FUNCTION_BLOCK FB_ModeSelect
VAR_INPUT
	bInterlockBypass: BOOL;
	bAutoPlayEnable: BOOL:=TRUE;
	sModuleDescription: STRING:='Mode Select';
	eModeZone:E_ModeZone;
	bLockedFB: BOOL;
	bPistonCheck: BOOL:=TRUE;
	bStateSafe_mode: BOOL:=TRUE;
END_VAR
VAR_OUTPUT
	bModeStillState: BOOL;
	bLockRequest: BOOL;
END_VAR
VAR
	fbPrintErrMessageByID: FB_PrintErrMessageByID_SFC_Cycle;
	r_trig_ModeExchange1: R_TRIG;
	r_trig_ModeExchange2: R_TRIG;
	r_trig_ModeExchange3: R_TRIG;
	ton_ModeExchengeDelay: TON;	
	fbOperation:FB_Operation;
	bLockRelay: BOOL;	
	i: INT;
	bPistonsOK: BOOL;
	fbFormatString:FB_FormatString;
	sFB_ID: STRING(3):='050';

	sActErrorID: STRING(11);
	sFullErrorId: STRING(11);
	//r_trigAuto: R_TRIG;
	r_trigIntClose: R_TRIG;
	r_trigIntOpen: R_TRIG;
	bIntZonePaused: BOOL;
	rt_Play: R_TRIG;

END_VAR
VAR
	ton_ResumeMachine: TON;
	ton_ResetErrors: TON;
	ton_ResetAllCycles: TON;
	ton_PlayAllDelay: TON;
	ton_PauseDelay: TON;
	r_trigPlayAllDelay: R_TRIG;
	ton_PlayDelay: TON;
END_VAR
VAR_IN_OUT
	stMode:ST_Mode;
	stOperation:ST_OperationButtons;
END_VAR

act_Oper();
act_ModeStillState();
fbOperation(stOper:=stOperation);
stMode.eModeZone:=eModeZone;		
stOperation.eModeZone:=eModeZone;
stOperation.sModeZone:=TO_STRING(eModeZone);
IF (stMode.iActMode=E_WorkingMode.eAutoMode OR stMode.iActMode=E_WorkingMode.eSemiAutoMode)
AND NOT bInterlockBypass
THEN;
	bLockRequest:=TRUE;
ELSE;
	bLockRequest:=FALSE;
END_IF



r_trigIntClose(CLK:=bLockedFB);
r_trigIntOpen(CLK:=NOT bLockedFB);

(*888888888888888888   InterLocks Zone 1		8888888888888*)
IF stOperation.iActOperation=E_OperationButtons.ePlayAll AND  r_trigIntOpen.Q THEN
	bIntZonePaused:=TRUE;
END_IF

IF NOT bLockedFB 
AND NOT bInterlockBypass	
AND stOperation.iActOperation=E_OperationButtons.ePlayAll THEN
	//Message
	sActErrorID:='351'; // '050x000x351',	'Warning',	'Interlock Paused Operation',
	act_GetErrorID_Format();
	fbPrintErrMessageByID(sFB_ModuleDescription:=sModuleDescription,sActErrorID:=sFullErrorId,bSFCError:=TRUE);
	stOperation.bSetPause:=TRUE;
	stOperation.iPauseHistory:=4;
END_IF


IF bAutoPlayEnable AND bIntZonePaused AND r_trigIntClose.Q THEN
	stOperation.bSetPlay:=TRUE;
	bIntZonePaused:=FALSE;
END_IF

IF bLockedFB OR stMode.iActMode=E_WorkingMode.eManualMode THEN
	bIntZonePaused:=FALSE;
END_IF

rt_Play(CLK:=stOperation.iActOperation=E_OperationButtons.ePlayAll);

IF NOT bStateSafe_mode OR stOperation.bStopResetAll THEN;
	stMode.bSetManual:=TRUE;
	stOperation.bSetPause:=TRUE;
END_IF

stMode.bStateSafe_mode:=stOperation.bStateSafe_mode:=bStateSafe_mode;

m_Error_zone_check();

stOperation.iActModeState:=stMode.iActMode;

ACTION act_AutomationLock_Failed:
sActErrorID:='306';//'050x000x306',	'Warning',	'Semi/Auto mode request rejected, automation lock failed',
act_GetErrorID_Format();
fbPrintErrMessageByID(sFB_ModuleDescription:=sModuleDescription,sActErrorID:=sFullErrorId,bSFCError:=TRUE);
END_ACTION

ACTION act_Done:
stMode.bSetManual:=FALSE;
stMode.bSetSemi:=FALSE;
stMode.bSetAuto:=FALSE;
//stMode.iErrorNum:=0;
//stMode.sErrorMessage:='No Error';
END_ACTION

ACTION act_GetErrorID_Format:
(*IF bErrorSFC THEN;
	
	IF    sLast_SFCErrorStep='WaitSenOpen' 							THEN sActErrorID:='001';
	ELSIF sLast_SFCErrorStep='WaitSenNotClose' 		   				THEN sActErrorID:='002';
	ELSIF sLast_SFCErrorStep='WaitSenClose' 						THEN sActErrorID:='003';
	ELSIF sLast_SFCErrorStep='WaitSenNotOpen' 						THEN sActErrorID:='004';
	ELSIF sLast_SFCErrorStep='No Status' 							THEN sActErrorID:='005';		
	ELSIF sLast_SFCErrorStep='No Valve Operation' 					THEN sActErrorID:='006';
	ELSIF sLast_SFCErrorStep='Not synchronized with cycle command' 	THEN sActErrorID:='007';
	ELSIF sLast_SFCErrorStep='SensorsChecking' 						THEN sActErrorID:='008';
	
	ELSE;
		 sActErrorID:='999';
	END_IF

ELSE
		 sActErrorID:='000';
END_IF*)

fbFormatString(
	sFormat:= '%.3sx%.3dx%.3s', 
	arg1:= F_STRINGEx(sFB_ID), 
	arg2:= F_INT(eModeZone), 
	arg3:= F_STRINGEx(sActErrorID), 
	sOut=>sFullErrorId );
END_ACTION

ACTION act_ModeStillState:

r_trig_ModeExchange1(CLK:=stMode.iActMode=eManualMode);
r_trig_ModeExchange2(CLK:=stMode.iActMode=eSemiAutoMode);
r_trig_ModeExchange3(CLK:=stMode.iActMode=eAutoMode);
ton_ModeExchengeDelay(PT:=T#0.5S);
(*IF ton_ModeExchengeDelay.Q THEN
	ton_ModeExchengeDelay.IN:=FALSE;
END_IF*)
IF r_trig_ModeExchange1.Q
OR r_trig_ModeExchange2.Q
OR r_trig_ModeExchange3.Q
THEN
	ton_ModeExchengeDelay(IN:=FALSE);
	ton_ModeExchengeDelay.IN:=TRUE;
END_IF
bModeStillState:=ton_ModeExchengeDelay.Q;
END_ACTION

ACTION act_Oper:
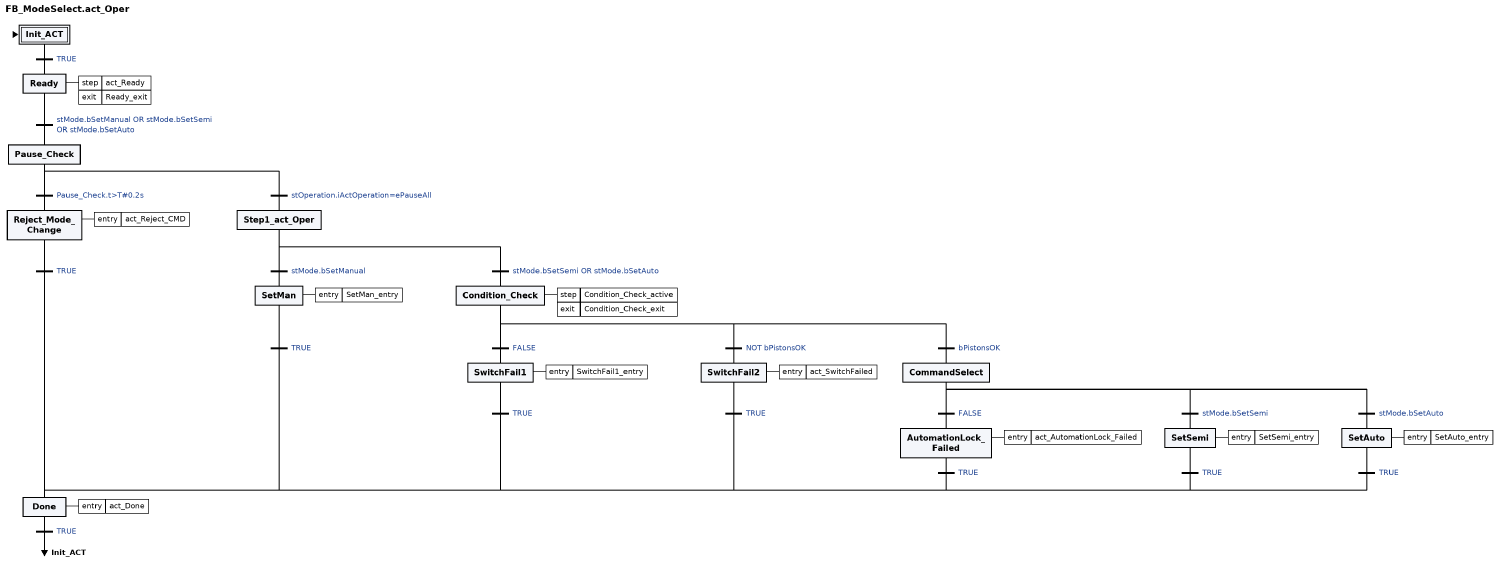
INITIAL_STEP Init_ACT:
END_STEP
TRANSITION FROM Init_ACT TO Ready
    := TRUE;
END_TRANSITION
STEP Ready:
    act_Ready(N);  // step action
    Ready_exit(P0);  // exit action
END_STEP
TRANSITION FROM Ready TO Pause_Check
    := stMode.bSetManual OR stMode.bSetSemi OR stMode.bSetAuto;
END_TRANSITION
STEP Pause_Check:
END_STEP
TRANSITION FROM Pause_Check TO Reject_Mode_Change
    := Pause_Check.t>T#0.2s;
END_TRANSITION
STEP Reject_Mode_Change:
    act_Reject_CMD(P1);  // entry action
END_STEP
TRANSITION FROM Reject_Mode_Change TO Done
    := TRUE;
END_TRANSITION
TRANSITION FROM Pause_Check TO Step1_act_Oper
    := stOperation.iActOperation=ePauseAll;
END_TRANSITION
STEP Step1_act_Oper:
END_STEP
TRANSITION FROM Step1_act_Oper TO SetMan
    := stMode.bSetManual;
END_TRANSITION
STEP SetMan:
    SetMan_entry(P1);  // entry action
END_STEP
TRANSITION FROM SetMan TO Done
    := TRUE;
END_TRANSITION
TRANSITION FROM Step1_act_Oper TO Condition_Check
    := stMode.bSetSemi OR stMode.bSetAuto;
END_TRANSITION
STEP Condition_Check:  // max time T#1s
    Condition_Check_active(N);  // step action
    Condition_Check_exit(P0);  // exit action
END_STEP
TRANSITION FROM Condition_Check TO SwitchFail1
    := FALSE;
END_TRANSITION
STEP SwitchFail1:
    SwitchFail1_entry(P1);  // entry action
END_STEP
TRANSITION FROM SwitchFail1 TO Done
    := TRUE;
END_TRANSITION
TRANSITION FROM Condition_Check TO SwitchFail2
    := NOT bPistonsOK;
END_TRANSITION
STEP SwitchFail2:
    act_SwitchFailed(P1);  // entry action
END_STEP
TRANSITION FROM SwitchFail2 TO Done
    := TRUE;
END_TRANSITION
TRANSITION FROM Condition_Check TO CommandSelect
    := bPistonsOK;
END_TRANSITION
STEP CommandSelect:  // max time T#1s
END_STEP
TRANSITION FROM CommandSelect TO AutomationLock_Failed
    := FALSE;
END_TRANSITION
STEP AutomationLock_Failed:
    act_AutomationLock_Failed(P1);  // entry action
END_STEP
TRANSITION FROM AutomationLock_Failed TO Done
    := TRUE;
END_TRANSITION
TRANSITION FROM CommandSelect TO SetSemi
    := stMode.bSetSemi;
END_TRANSITION
STEP SetSemi:
    SetSemi_entry(P1);  // entry action
END_STEP
TRANSITION FROM SetSemi TO Done
    := TRUE;
END_TRANSITION
TRANSITION FROM CommandSelect TO SetAuto
    := stMode.bSetAuto;
END_TRANSITION
STEP SetAuto:
    SetAuto_entry(P1);  // entry action
END_STEP
TRANSITION FROM SetAuto TO Done
    := TRUE;
END_TRANSITION
STEP Done:
    act_Done(P1);  // entry action
END_STEP
TRANSITION FROM Done TO Init_ACT
    := TRUE;
END_TRANSITION
// branch label Branch3_act_Oper
// branch label Branch1_act_Oper
// branch label Branch0_ACT
// branch label Branch2_act_Oper
END_ACTION

ACTION act_Operation:
(*
IF stOperation.bSetPlay THEN;
	bResumeMachine:=TRUE;
END_IF
ton_ResumeMachine(PT:=T#10MS,IN:=bResumeMachine,);
ton_PlayAllDelay(PT:=T#20MS);
IF ton_ResumeMachine.Q THEN;
	bResumeMachine:=FALSE;	
	stOperation.bSetPlay:=FALSE;
	ton_PlayAllDelay.IN:=TRUE;	
END_IF





r_trigPlayAllDelay(CLK:=ton_PlayAllDelay.Q);
IF r_trigPlayAllDelay.Q THEN	
	IF FALSE(*iActErrorNum=0*) THEN
		//stOperation.iActOperation:=E_OperationButtons.ePlayAll;
		stOperation.bSetPlay:=TRUE;
	END_IF	
END_IF


IF stOperation.bSetPause THEN;
	stOperation.iActOperation:=E_OperationButtons.ePauseAll;
	stOperation.bSetPause:=FALSE;
	ton_PlayAllDelay.IN:=FALSE;
END_IF



IF stOperation.iActOperation=E_OperationButtons.ePauseAll THEN;
	
ELSIF stOperation.iActOperation=E_OperationButtons.ePlayAll THEN;
	
END_IF

bPauseMachine:=stOperation.iActOperation=E_OperationButtons.ePauseAll;


ton_PauseDelay(PT:=T#1S, IN:=stOperation.iActOperation=E_OperationButtons.ePauseAll);
ton_PlayDelay(PT:=T#1S, IN:=stOperation.iActOperation=E_OperationButtons.ePlayAll);
*)
END_ACTION

ACTION act_Ready:

IF stMode.iActMode=eManualMode AND stMode.bSetManual THEN; stMode.bSetManual:=FALSE; END_IF
IF stMode.iActMode=eSemiAutoMode AND stMode.bSetSemi THEN; stMode.bSetSemi:=FALSE; END_IF

IF stMode.iActMode=eAutoMode 
AND stMode.bSetAuto THEN; 
	stMode.bSetAuto:=FALSE; 
ELSIF stMode.iActMode=eAutoMode 
AND stMode.bSetSemi THEN; 
	stMode.bSetSemi:=FALSE;	
	stMode.iActMode:=eSemiAutoMode;
END_IF

IF stOperation.bStopResetAll THEN;
	stMode.bSetManual:=TRUE;
END_IF
END_ACTION

ACTION act_Reject_CMD:

	IF stMode.bSetManual 	THEN; sActErrorID:='300';END_IF	(*	'050x000x300',	'Warning',	'Manual mode request rejected, first pause automation',	*)
	IF stMode.bSetSemi 		THEN; sActErrorID:='301';END_IF	(*	'050x000x301',	'Warning',	'Semi mode request rejected, first pause automation',	*)
	IF stMode.bSetAuto 		THEN; sActErrorID:='302';END_IF	(*	'050x000x302',	'Warning',	'Auto mode request rejected, first pause automation',	*)
	act_GetErrorID_Format();
	fbPrintErrMessageByID(sFB_ModuleDescription:=sModuleDescription,sActErrorID:=sFullErrorId,bSFCError:=TRUE);
END_ACTION

ACTION act_SwitchFailed:

IF stMode.bSetManual 	THEN; sActErrorID:='303';END_IF	(*	'050x000x303',	'Warning',	'Manual mode request rejected, Pistion not in last auto pisition',	*)
IF stMode.bSetSemi 		THEN; sActErrorID:='304';END_IF	(*	'050x000x304',	'Warning',	'Semi mode request rejected, Pistion not in last auto pisition',	*)
IF stMode.bSetAuto 		THEN; sActErrorID:='304';END_IF	(*	'050x000x305',	'Warning',	'Auto mode request rejected, Pistion not in last auto pisition',	*)
act_GetErrorID_Format();
fbPrintErrMessageByID(sFB_ModuleDescription:=sModuleDescription,sActErrorID:=sFullErrorId,bSFCError:=TRUE);

stMode.bSetManual:=FALSE;
stMode.bSetSemi:=FALSE;
stMode.bSetAuto:=FALSE;
END_ACTION

ACTION Condition_Check_active:
bPistonsOK:=TRUE;
IF bPistonCheck THEN
	FOR i:=1 TO C_Max_Pistons DO;
		IF stPis[i].b_Exist
		AND (NOT stPis[i].st_SyncAuto) THEN;
			IF stPis[i].eModeZone=eModeZone THEN;
				stPis[i].b_Print_NotSyncAutoMessage:=TRUE;
				bPistonsOK:=FALSE;
			END_IF
		END_IF
	END_FOR	
END_IF
END_ACTION

ACTION Condition_Check_exit:
IF NOT bPistonsOK THEN;	
(*	IF stMode.bSetManual 	THEN; sActErrorID:='303';END_IF	(*	'050x000x303',	'Warning',	'Manual mode request rejected, Pistion not in last auto pisition',	*)
	IF stMode.bSetSemi 		THEN; sActErrorID:='304';END_IF	(*	'050x000x304',	'Warning',	'Semi mode request rejected, Pistion not in last auto pisition',	*)
	IF stMode.bSetAuto 		THEN; sActErrorID:='304';END_IF	(*	'050x000x305',	'Warning',	'Auto mode request rejected, Pistion not in last auto pisition',	*)
	act_GetErrorID_Format();
	fbPrintErrMessageByID(sModuleDescription:=sModuleDescription,sActErrorID:=sFullErrorId);*)
END_IF
END_ACTION

METHOD m_Error_zone_check : BOOL
VAR_INPUT
END_VAR

VAR
	i: INT;
	sCheckZone: STRING;

END_VAR
sCheckZone:=TO_STRING(stMode.eModeZone);

FOR i:=1 TO C_Max_Buffer_Act_list DO;
	IF TRUE 
	AND Buffer_Act_Message[i].sLevel='Error'
	AND Buffer_Act_Message[i].sModuleDescription=sCheckZone
	AND stOperation.iActOperation=E_OperationButtons.ePlayAll 
	THEN;
		stOperation.bSetPause:=TRUE;
	END_IF
END_FOR
END_METHOD

ACTION Ready_exit:
stOperation.bSetPause:=TRUE;
stOperation.iPauseHistory:=6;
END_ACTION

ACTION SetAuto_entry:
stMode.iActMode:=eAutoMode;
END_ACTION

ACTION SetMan_entry:
stMode.iActMode:=eManualMode;
END_ACTION

ACTION SetSemi_entry:
stMode.iActMode:=eSemiAutoMode;
END_ACTION

ACTION SwitchFail1_entry:
//entrance condition <NOT prg_Initialise.bGeneralDone>

//IF stMode.bSetAuto 		THEN; sActErrorID:='304';END_IF	(*	'050x000x305',	'Warning',	'Auto mode request rejected, Pistion not in last auto pisition',	*)

sActErrorID:='350'; // '050x000x350',	'Warning',	'Semi/Auto mode request rejected, initialize all system first',
act_GetErrorID_Format();
fbPrintErrMessageByID(sFB_ModuleDescription:=sModuleDescription,sActErrorID:=sFullErrorId,bSFCError:=TRUE);

stMode.bSetManual:=FALSE;
stMode.bSetSemi:=FALSE;
stMode.bSetAuto:=FALSE;
END_ACTION

END_FUNCTION_BLOCK

(* stored: Version 1.1.0.1, ProductVersion 3.1.4024.13
   POU FB_ModeSelect: Id {b95347f3-88f5-4be2-b47c-79ac89a3355f}, SpecialFunc None
   Folder Actions: Id {82255ca1-1f75-456a-a29d-0d95ddaf34af}
   Action act_AutomationLock_Failed: Id {749ee08a-32c4-42e6-baa7-e0e1eee12535}
   Action act_Done: Id {296eb8e7-61ec-4e1e-9dc0-d90c1d2d741e}
   Action act_GetErrorID_Format: Id {06fa01f5-e787-4c81-a2b4-ad12d608a7c8}
   Action act_ModeStillState: Id {8ed3c8be-df69-41c3-95fa-f76f61afeb74}
   Action act_Oper: Id {e7dcf637-733d-4980-abb2-53e9ba8fbeff}
   Action act_Operation: Id {d99501f7-9523-4197-a4a8-8762849e15ea}
   Action act_Ready: Id {0b6aadda-085e-4ced-978e-c2e348c4875f}
   Action act_Reject_CMD: Id {29be06db-0135-4037-bf95-33eaa49632e7}
   Action act_SwitchFailed: Id {0bafcad7-61fd-48ec-8730-f5aebd8fa624}
   Action Condition_Check_active: Id {e128942e-0ef4-40fb-bfd1-9a6e83cafa0d}
   Action Condition_Check_exit: Id {71572210-e632-4875-9651-3697c7764c07}
   Method m_Error_zone_check: Id {d71a2d60-edec-4d86-b797-3285b49c2480}
   Action Ready_exit: Id {ab53e8f1-23f1-4ef5-9d62-59ff46d788ce}
   Action SetAuto_entry: Id {906f77fe-e6af-4363-a7f2-9a8ea55499dc}
   Action SetMan_entry: Id {35c0470c-3ef9-4a62-a98e-99801a1845c6}
   Action SetSemi_entry: Id {d2dffbfe-e7bb-4d4a-81f3-bbc52c51799f}
   Action SwitchFail1_entry: Id {0a54deee-f1fc-4dfc-972d-717bcd92630a} *)
